// TIA Portal V20 export
// export: Created 2026-10-12T04:58:20.6627774Z, ExportSetting WithDefaults, DisplayName Totally Integrated Automation Portal, DisplayVersion V20, DisplayName TIA Portal Openness, DisplayVersion V20, DisplayName TIA Portal Teamcenter Gateway, DisplayVersion V20, DisplayName TIA Portal Version Control Interface, DisplayVersion V20, DisplayName SINAMICS Startdrive Advanced, DisplayVersion V20 SP1 Update 2, DisplayName SINAMICS Startdrive G110M, G120, G120C, G120D, G120P, G115D, DisplayVersion V20 SP1 Update 2, DisplayName SINAMICS Startdrive G130, G150, S120, S150, SINAMICS MV, G220, S200, S210, DisplayVersion V20 SP1 Update 2, DisplayName STEP 7 Professional, DisplayVersion V20, DisplayName STEP 7 Safety, DisplayVersion V20, DisplayName WinCC Basic/Comfort/Advanced, DisplayVersion V20, DisplayName WinCC Professional, DisplayVersion V20, DisplayName WinCC Unified, DisplayVersion V20
FUNCTION "FRK_UnitModeResolve" : Void   // FC74, SCL
{ S7_Optimized_Access := 'TRUE' }
VERSION : 0.1
// stored: AutoNumber true, IsIECCheckEnabled false, SetENOAutomatically false, UDAEnableTagReadback false
   VAR_INPUT
      Policy : Array[0..6] of "ST_ModePolicy";
      Timeout : Time;
   END_VAR
   VAR_IN_OUT
      Core : "FRK_Core";
      Unit : "FRK_Unit";
      Status : "ST_ModuleStatus";
   END_VAR
BEGIN

   IF #Unit.ModePending THEN
       IF #Timeout <= T#0ms OR "FRK_Elapsed"(NewMs := "FRK_Clock".NowMs, OldMs := #Unit.ModeSince) >= DINT_TO_UDINT(TIME_TO_DINT(#Timeout)) THEN
           "FRK_Fault"(Core := #Core,
                       Status := #Status,
                       ReasonCode := 2001,
                       Description := WSTRING#'std.error.hmiRequestRejected');
           #Unit.ModePending := FALSE;
           #Unit.FollowStart := FALSE;
           #Unit.ReleaseChildren := TRUE;
           #Unit.Clearing := TRUE;
       ELSIF #Core.EvModeExit THEN
           #Unit.ExitFirst := FALSE;
           IF #Policy[#Unit.Mode].Style = 0 THEN
               #Unit.StopReq := TRUE;
           ELSIF #Core.HookResult <= 0 THEN
               #Unit.AbortReq := TRUE;
               #Unit.ReleaseChildren := TRUE;
               #Unit.Clearing := TRUE;
           END_IF;
       END_IF;
   END_IF;
END_FUNCTION
